Staubli VAL3: resetOutput.pgx

public program resetOutput()
  local bool l_bErr
  local num l_nI
begin
  //2025.7.21 add 复位输出信号
  for l_nI=9 to size(io:dOutput)-1
    call io:setDigOutput(io:dOutput[l_nI],false,l_bErr)
  endFor
  for l_nI=0 to size(io:aOutput)-1
    call io:setAnaOutput(io:aOutput[l_nI],0,l_bErr)
  endFor
end
